FUNCTION_BLOCK SKILL_Core (* The part every skill shares: its state machine (Idle, Running, Stopping, Succeeded, Failed, Aborted), the OPC UA methods Stop, Abort and Reset, and the State and ErrorID it publishes. It checks a client's Start (the caller holds the occupation, the module is in Execute, the skill is not running, the values are in range, the equipment is free) and then starts the skill's own logic. Technical: Skill core: state machine, OPC UA Stop/Abort/Reset(Session) -> [Accepted, ErrorID], State and ErrorID published, activity counted; the Start method (with the skill's parameters) is wired to START_REQ and START_RSP; RUN starts the execution, SUCCESS or FAILURE(ErrorID) ends it *)
  (* Standard: 61499-2 *)
  (* Version 0.1, 2026-09-28, Project contributors, AAU Smart Production Lab *)
  PACKAGE modlib;
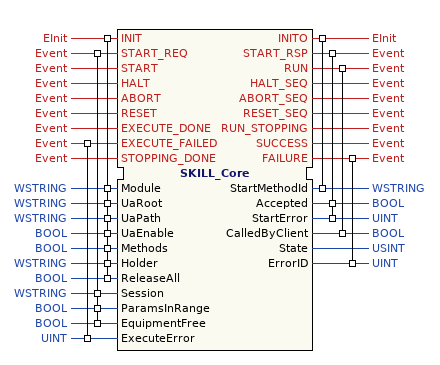
  EVENT_INPUT
    INIT : EInit WITH Module, UaRoot, UaPath, UaEnable, Methods, Holder, ReleaseAll; (* Initialise, once at start-up (the INIT chain); takes the values given with it *)
    START_REQ WITH Session, ParamsInRange, EquipmentFree; (* Start(Session, parameters) was called: check Session, ParamsInRange, EquipmentFree *)
    START; (* Start a run, from the parent (a step of a sequence): no session check *)
    HALT; (* Stop the run, from the parent *)
    ABORT; (* Abort: everything off at once *)
    RESET; (* Reset from Failed or Aborted to Idle *)
    EXECUTE_DONE; (* The execution ended successfully *)
    EXECUTE_FAILED WITH ExecuteError; (* The execution failed (ExecuteError) *)
    STOPPING_DONE; (* The stop sequence ended *)
  END_EVENT
  EVENT_OUTPUT
    INITO : EInit WITH StartMethodId; (* Initialised: the next block of the INIT chain goes on *)
    START_RSP WITH Accepted, StartError; (* Answer to Start *)
    RUN WITH CalledByClient; (* Run: latch the parameters, start the execution *)
    HALT_SEQ; (* Halt the execute sequence *)
    ABORT_SEQ; (* Abort the sequences *)
    RESET_SEQ; (* Reset the sequences *)
    RUN_STOPPING; (* Run the stop sequence (the skill was stopped) *)
    SUCCESS; (* The run succeeded (the results are set) *)
    FAILURE WITH ErrorID; (* The run failed (ErrorID) *)
  END_EVENT
  VAR_INPUT
    Module : WSTRING; (* The module's name; its local channels are named after it (loc[<Module>/...]) *)
    UaRoot : WSTRING; (* The module's OPC UA folder, e.g. /Objects/Filling *)
    UaPath : WSTRING; (* This skill's OPC UA folder below UaRoot, e.g. /Skills/Dispensing *)
    UaEnable : BOOL; (* Publish on OPC UA *)
    Methods : BOOL; (* Offer the OPC UA methods Start, Stop, Abort, Reset (FALSE: a step, run by its parent) *)
    Holder : WSTRING; (* The name the equipment is held under: the skill's own, or for a step the skill it belongs to *)
    ReleaseAll : BOOL := FALSE; (* When a run ends, give up everything held under Holder (a module level skill) *)
    Session : WSTRING; (* Session ID of the caller of Start (must be the module's owner) *)
    ParamsInRange : BOOL := TRUE; (* Every Start argument lies within its limits *)
    EquipmentFree : BOOL := TRUE; (* The equipment is free, or held by this skill *)
    ExecuteError : UINT; (* Why the execution failed *)
  END_VAR
  VAR_OUTPUT
    StartMethodId : WSTRING; (* OPC UA ID of the Start method, for its SERVER block *)
    Accepted : BOOL; (* The call was accepted *)
    StartError : UINT; (* Why Start was refused (error code) *)
    CalledByClient : BOOL; (* Started over OPC UA (take the Start arguments), not by a parent (take the defaults) *)
    State : USINT; (* Skill state: 0 Idle, 1 Running, 2 Stopping, 3 Succeeded, 4 Failed, 5 Aborted *)
    ErrorID : UINT; (* Error code: 0 none, 1 PreconditionViolated, 2 InvariantViolated, 3 Timeout, 4 NotReady, 5 NotPermitted, 6 Busy, 7 Interrupted, 8 OutOfRange *)
  END_VAR
  (* Group StateMachine: The skill's states; in front of them the gate, which decides a client's command; and when a Succeeded returns to Idle *)
  (* Group ModuleViews: The module's owner and state in, the activity count out *)
  (* Group OpcUa: The methods Stop, Abort and Reset, and the published State and ErrorID *)
  (* Group Release: At the end of a run of a module level skill: everything it holds given up *)
  FBS
    Gate : modlib::SKILL_Gate; (* Decides a client's Start, Stop, Abort and Reset and answers it; passes accepted ones, and the parent's commands, on to Control. *) {SET_ATTRIBUTE(GroupName, StateMachine)}
    Control : modlib::SKILL_Control; (* The skill's state machine (SKILL_Control). *) {SET_ATTRIBUTE(GroupName, StateMachine)}
    Owner : modlib::MOD_OwnerView; (* Knows who occupies the module: only the owner may command the skill over OPC UA. *) {SET_ATTRIBUTE(GroupName, ModuleViews)}
    Mode : modlib::MOD_StateView; (* Knows the module's state: a client may start the skill only in Execute; the skill stops when the module stops. *) {SET_ATTRIBUTE(GroupName, ModuleViews)}
    UaStop : iec61499::net::SERVER_2_1; (* The OPC UA method Stop(Session). *) {SET_ATTRIBUTE(GroupName, OpcUa)}
    UaAbort : iec61499::net::SERVER_2_1; (* The OPC UA method Abort(Session). *) {SET_ATTRIBUTE(GroupName, OpcUa)}
    UaReset : iec61499::net::SERVER_2_1; (* The OPC UA method Reset(Session). *) {SET_ATTRIBUTE(GroupName, OpcUa)}
    PubState : iec61499::net::PUBLISH_2; (* Writes State and ErrorID to OPC UA. *) {SET_ATTRIBUTE(GroupName, OpcUa)}
    Act : iec61499::net::PUBLISH_1(QI := TRUE); (* Says +1 when the skill starts and -1 when it ends, for the module's count of running skills. *) {SET_ATTRIBUTE(GroupName, ModuleViews)}
    ToIdle : iec61499::events::E_DELAY(DT := T#1500ms); (* Brings a succeeded skill back to Idle after 1.5 s. *) {SET_ATTRIBUTE(GroupName, StateMachine)}
    PubRelease : iec61499::net::PUBLISH_1; (* When a run ends, says on the release channel that this skill gives up its equipment. *) {SET_ATTRIBUTE(GroupName, Release)}
  END_FBS
  EVENT_CONNECTIONS
    INIT TO Control.INIT;
    Control.INITO TO Owner.INIT;
    Owner.INITO TO Mode.INIT;
    Mode.INITO TO UaStop.INIT;
    UaStop.INITO TO UaAbort.INIT;
    UaAbort.INITO TO UaReset.INIT;
    UaReset.INITO TO PubState.INIT;
    PubState.INITO TO Act.INIT;
    Act.INITO TO PubRelease.INIT;
    PubRelease.INITO TO PubState.REQ;
    PubRelease.INITO TO INITO;
    START_REQ TO Gate.START_REQ;
    Gate.START_RSP TO START_RSP;
    UaStop.IND TO Gate.STOP_REQ;
    Gate.STOP_RSP TO UaStop.RSP;
    UaAbort.IND TO Gate.ABORT_REQ;
    Gate.ABORT_RSP TO UaAbort.RSP;
    UaReset.IND TO Gate.RESET_REQ;
    Gate.RESET_RSP TO UaReset.RSP;
    Owner.CHG TO Gate.OWNER_CHG;
    Mode.CHG TO Gate.MOD_CHG;
    Gate.GO_START TO Control.START;
    Gate.GO_HALT TO Control.HALT;
    Gate.GO_ABORT TO Control.ABORT;
    Gate.GO_RESET TO Control.RESET;
    Control.PUB TO PubState.REQ;
    Control.PUB TO Gate.SKILL_CHG;
    Control.ACT TO Act.REQ;
    START TO Gate.START;
    HALT TO Gate.HALT;
    ABORT TO Gate.ABORT;
    RESET TO Gate.RESET;
    EXECUTE_DONE TO Control.EXECUTE_DONE;
    EXECUTE_FAILED TO Control.EXECUTE_FAILED;
    STOPPING_DONE TO Control.STOPPING_DONE;
    Control.RUN TO RUN;
    Control.HALT_SEQ TO HALT_SEQ;
    Control.ABORT_SEQ TO ABORT_SEQ;
    Control.RESET_SEQ TO RESET_SEQ;
    Control.RUN_STOPPING TO RUN_STOPPING;
    Control.SUCCESS TO SUCCESS;
    Control.FAILURE TO FAILURE;
    Control.TO_IDLE_START TO ToIdle.START;
    Control.TO_IDLE_STOP TO ToIdle.STOP;
    ToIdle.EO TO Control.TO_IDLE;
    Control.RELEASE TO PubRelease.REQ;
  END_CONNECTIONS
  DATA_CONNECTIONS
    Module TO Control.Module;
    Module TO Owner.Module;
    Module TO Mode.Module;
    UaRoot TO Control.UaRoot;
    UaPath TO Control.UaPath;
    Methods TO UaStop.QI;
    Methods TO UaAbort.QI;
    Methods TO UaReset.QI;
    UaEnable TO PubState.QI;
    Control.StartMethodId TO StartMethodId;
    Session TO Gate.Session;
    ParamsInRange TO Gate.ParamsInRange;
    EquipmentFree TO Gate.EquipmentFree;
    Gate.Accepted TO Accepted;
    Gate.Accepted TO UaStop.SD_1;
    Gate.Accepted TO UaAbort.SD_1;
    Gate.Accepted TO UaReset.SD_1;
    Gate.ResponseError TO StartError;
    Gate.ResponseError TO UaStop.SD_2;
    Gate.ResponseError TO UaAbort.SD_2;
    Gate.ResponseError TO UaReset.SD_2;
    Control.StopMethodId TO UaStop.ID;
    UaStop.RD_1 TO Gate.StopSession;
    Control.AbortMethodId TO UaAbort.ID;
    UaAbort.RD_1 TO Gate.AbortSession;
    Control.ResetMethodId TO UaReset.ID;
    UaReset.RD_1 TO Gate.ResetSession;
    Owner.Owner TO Gate.Owner;
    Mode.State TO Gate.ModuleState;
    Gate.ByClient TO Control.ByClient;
    Control.StateId TO PubState.ID;
    Control.State TO PubState.SD_1;
    Control.State TO State;
    Control.State TO Gate.State;
    Control.ErrorID TO PubState.SD_2;
    Control.ErrorID TO ErrorID;
    Control.ActivityId TO Act.ID;
    Control.ActivityDelta TO Act.SD_1;
    ExecuteError TO Control.ExecuteError;
    Control.CalledByClient TO CalledByClient;
    ReleaseAll TO PubRelease.QI;
    Control.ReleaseId TO PubRelease.ID;
    Holder TO PubRelease.SD_1;
  END_CONNECTIONS
END_FUNCTION_BLOCK
